(* IEC 61131-3 sources: openplc-editor-canopen/e2e/fixtures/canopen-boot-sdo/project/pous/programs, 1 file *)

(* ---- main.st ---- *)
PROGRAM main
  VAR
    inputs AT %IB1 : BYTE;
    outputs AT %QB0 : BYTE;
  END_VAR

outputs := inputs;

END_PROGRAM
